Staubli VAL3: main.pgx

program main()
begin
  close(tCurrentTool)
  pPointRx.config.shoulder = lefty
  pPointRx.config.elbow = epositive
  pPointRx.config.wrist = wpositive
  pPointRx2.config.shoulder = lefty
  pPointRx2.config.elbow = epositive
  pPointRx2.config.wrist = wpositive
  mCurrentSpeed.tvel = 100.00
  mCurrentSpeed.blend = joint
  mCurrentSpeed.reach = 0.010
  mCurrentSpeed.leave = 0.010
  // Program EdgeProg start
  // Program generated by RoboDK v6.0.7 for Staubli RX130B on XX/XX/XXXX 18:00:00
  // Using nominal kinematics.
  mCurrentSpeed.tvel = 123.456
  mCurrentSpeed.reach = -1.000
  mCurrentSpeed.leave = -1.000
  call MoveJoint(-5.00000,-5.00000,15.00000,10.00000,40.00000,-10.00000)
  mCurrentSpeed.reach = 12.500
  mCurrentSpeed.leave = 12.500
  pPointRx.config.wrist = wnegative
  call MoveLine(-624.230,571.208,454.620,81.604,51.756,-128.588)
  delay(0.000)
  delay(1.234)
  popUpMsg("A long message with "quotes", 'apostrophes' & symbols: <>[]{}()=+-*/%;#@! and more text to make it longer than eighty characters")
  // Comment with ; semicolon
  Gripper=ON
  Output[12]=false
  Pressure=true
  watch(PartPresent==true,250.0)
  watch(Input[7]==1)
  //call prog:Do Something(1, 2)
  x = 1
  call MoveJoint(20.00000,-10.00000,20.00000,0.00000,30.00000,0.00000)

  waitEndMove()
  // Program EdgeProg end

end
